Fanuc KAREL source: KA00016.KL

PROGRAM KA00016
%NOLOCKGROUP
VAR
  SRC: REAL
  DST: STRING[80]
BEGIN
  SRC = 2.0
  DST = SRC
END KA00016
